SUBAPPLICATION Uebung_146 (* Übung zu RATE: Wiederholrate 1000/100 ms zur Laufzeit (Grenzen 50..2000 ms) *)
  (* Standard: 61499-2; Description: Copyright (c) 2023 Meisterschulen am Ostbahnhof This program and the accompanying materials are made available under the terms of the Eclipse Public License 2.0 which is available at https://www.eclipse.org/legal/epl-2.0/ SPDX-License-Identifier: EPL-2.0 *)
  (* Version 1.0, 2026-11-17, Franz Höpfinger, Meisterschulen am Ostbahnhof, initial API and implementation and/or initial documentation *)
  PACKAGE Uebungen;
  IMPORT Uebungen::const::Uebung_120_129::Filter::PEAK_ADD;
  IMPORT Uebungen::const::Uebung_120_129::Filter::PEAK_FLT;
  IMPORT isobus::pgn::ISOUSERHOME_e::network;
  IMPORT isobus::pgn::ISO_CAN_NODE::NODE1;
  IMPORT isobus::pgn::const::PgnDef::PGN_PDU1_PropA;
  IMPORT logiBUS::io::DI::logiBUS_DI::Input_I2;
  IMPORT logiBUS::io::DI::logiBUS_DI_Events::BUTTON_SINGLE_CLICK;
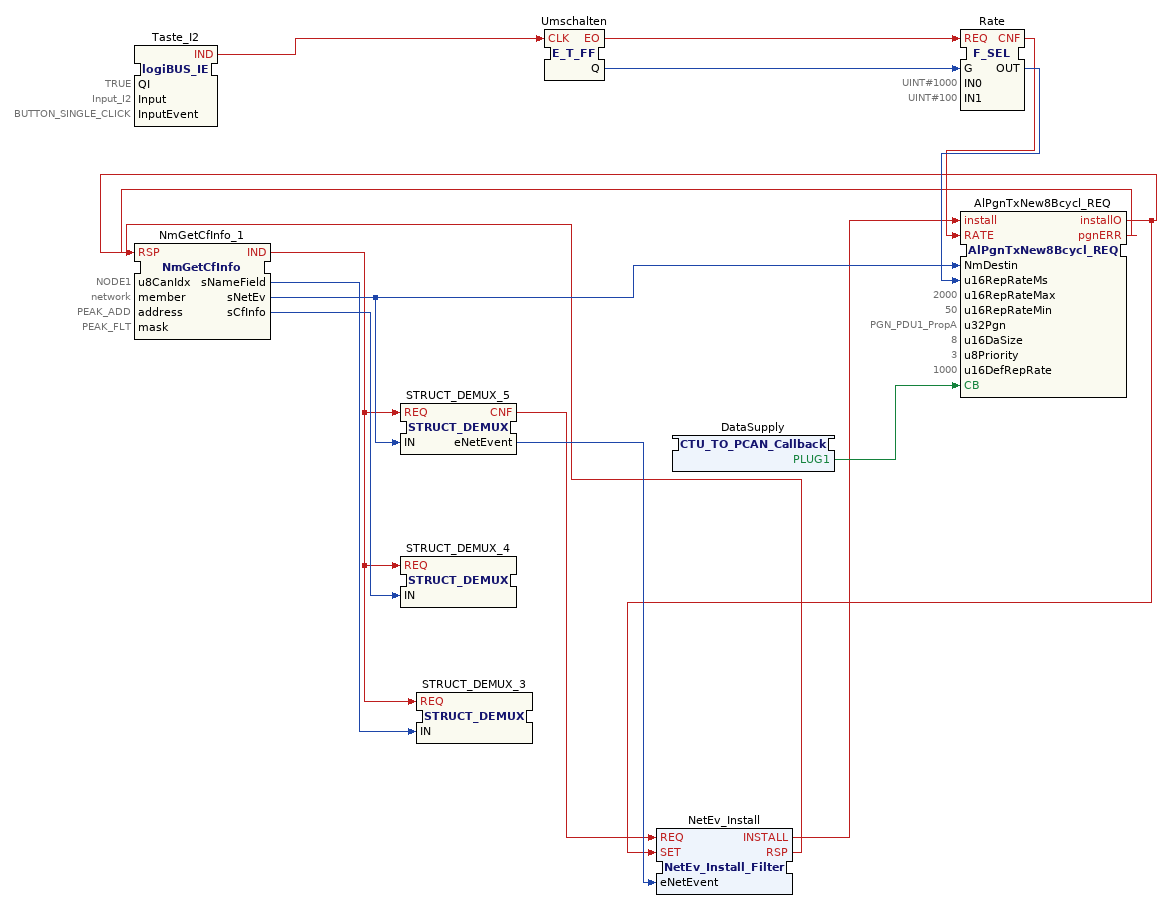
  (* RATE: Wiederholrate zur Laufzeit ändern (AlPgnTxNew8Bcycl_REQ) Grenzen beim install: u16RepRateMin 50, u16RepRateMax 2000 ms (beide ungleich 0, sonst RATE = pgnERR E_CONFIG). Start 1000 ms. I2 Klick: 100 ms, nochmal: 1000 ms. Außerhalb 50..2000: pgnERR E_VALUE_WRONG. *)
  FBS
    STRUCT_DEMUX_3 : eclipse4diac::convert::STRUCT_DEMUX; {SET_ATTRIBUTE(StructuredType, isobus::pgn::NAMEFIELD_T)}
    NmGetCfInfo_1 : isobus::pgn::NmGetCfInfo(u8CanIdx := NODE1, member := network, address := PEAK_ADD, mask := PEAK_FLT);
    STRUCT_DEMUX_4 : eclipse4diac::convert::STRUCT_DEMUX; {SET_ATTRIBUTE(StructuredType, isobus::pgn::CF_INFO_T)}
    STRUCT_DEMUX_5 : eclipse4diac::convert::STRUCT_DEMUX; {SET_ATTRIBUTE(StructuredType, isobus::pgn::ISONETEVENT_T)}
    AlPgnTxNew8Bcycl_REQ : isobus::pgn::tx::AlPgnTxNew8Bcycl_REQ(u16RepRateMax := 2000, u16RepRateMin := 50, u32Pgn := PGN_PDU1_PropA, u16DaSize := 8, u8Priority := 3, u16DefRepRate := 1000);
    Taste_I2 : logiBUS::io::DI::logiBUS_IE(QI := TRUE, Input := Input_I2, InputEvent := BUTTON_SINGLE_CLICK);
    Umschalten : iec61499::events::E_T_FF;
    Rate : iec61131::selection::F_SEL(IN0 := UINT#1000, IN1 := UINT#100); (* Q=FALSE: 1000 ms, Q=TRUE: 100 ms *)
  END_FBS
  SUBAPPS
    DataSupply : MyLib::sys::CTU_TO_PCAN_Callback;
    NetEv_Install : MyLib::sys::NetEv_Install_Filter;
  END_SUBAPPS
  EVENT_CONNECTIONS
    NmGetCfInfo_1.IND TO STRUCT_DEMUX_3.REQ;
    NmGetCfInfo_1.IND TO STRUCT_DEMUX_4.REQ;
    NmGetCfInfo_1.IND TO STRUCT_DEMUX_5.REQ;
    AlPgnTxNew8Bcycl_REQ.installO TO NmGetCfInfo_1.RSP;
    AlPgnTxNew8Bcycl_REQ.pgnERR TO NmGetCfInfo_1.RSP;
    STRUCT_DEMUX_5.CNF TO NetEv_Install.REQ;
    NetEv_Install.INSTALL TO AlPgnTxNew8Bcycl_REQ.install;
    NetEv_Install.RSP TO NmGetCfInfo_1.RSP;
    AlPgnTxNew8Bcycl_REQ.installO TO NetEv_Install.SET;
    Taste_I2.IND TO Umschalten.CLK;
    Umschalten.EO TO Rate.REQ;
    Rate.CNF TO AlPgnTxNew8Bcycl_REQ.RATE;
  END_CONNECTIONS
  DATA_CONNECTIONS
    NmGetCfInfo_1.sNameField TO STRUCT_DEMUX_3.IN;
    NmGetCfInfo_1.sNetEv TO STRUCT_DEMUX_5.IN;
    NmGetCfInfo_1.sCfInfo TO STRUCT_DEMUX_4.IN;
    NmGetCfInfo_1.sNetEv TO AlPgnTxNew8Bcycl_REQ.NmDestin;
    STRUCT_DEMUX_5.eNetEvent TO NetEv_Install.eNetEvent;
    Umschalten.Q TO Rate.G;
    Rate.OUT TO AlPgnTxNew8Bcycl_REQ.u16RepRateMs;
  END_CONNECTIONS
  ADAPTER_CONNECTIONS
    DataSupply.PLUG1 TO AlPgnTxNew8Bcycl_REQ.CB;
  END_CONNECTIONS
END_SUBAPPLICATION
